Fanuc KAREL source: KA00061.KL

PROGRAM KA00061
%NOLOCKGROUP
VAR
  SRC: XYZWPR
  DST: INTEGER
BEGIN
  SRC.X = 1.0
  DST = SRC
END KA00061
